TYPE ST_JointTarget :
STRUCT
	Position : ST_JointPose; // Commanded joint angles
    Velocity : ST_JointVelocity; // Commanded joint speeds
    Torque   : ST_JointTorque; // Calculated motor torques (T1, T2, T3)
END_STRUCT
END_TYPE

(* stored: Version 1.1.0.1, ProductVersion 3.1.4024.15
   DUT ST_JointTarget: Id {c381f50e-42a7-4e2e-889c-8b5a755635f1} *)
